Staubli VAL3: getTrajID.pgx

program getTrajID()
  local num l_nSession
  local num i
  local string l_sEmpty
  local bool l_bOk
begin
  // init
  //  x_bFounded=false
  //  x_sSessionName=""
  //  //
  // get the list
  //
  //  l_sEmpty=""
  call trajectory:getTrajList(sSessionList)
  //
  // search the program from a number:
  //
  // "number+space+name"
  //
  // 01 MyPart
  // 10 YourPart
  //
  resize(nIDIsExit,1,size(sSessionList))
  for i=0 to size(sSessionList)-1
    if sSessionList[i]!=""
      // convert the string "00 name" into a num
      toNum(sSessionList[i],l_nSession,l_bOk)
      if l_bOk
        nIDIsExit[i]=l_nSession
        endIf
    endIf
  endFor
end
